(*
SPDX-FileCopyrightText: © 2026 Oleksandr Tiutyk <trofimich@gmail.com>
SPDX-License-Identifier: MIT
License: https://opensource.org/license/mit
*)

(*!
<summary>
Defines a composite activity that waits until the first branch condition becomes TRUE and runs its activity.
</summary>
*)

INTERFACE IWaitAndPickActivity EXTENDS IExclusiveCompositeActivity

(*!
<summary>Appends a condition-activity branch pair and returns its zero-based branch index.</summary>
<description>
Permitted only in PASSIVE_READY. Both condition and activity are required and must not be attached elsewhere.
The standard implementation also rejects duplicate slots, validates fixed workflow association and requires
the parent chain and owning workflow to be PASSIVE_READY before mutation. Child storage remains borrowed.
</description>
<param name="condition">Condition evaluated when polling branches in registration order.</param>
<param name="activity">Activity executed once condition evaluates to TRUE.</param>
*)
METHOD AddBranch : DINT
VAR_INPUT
	condition : ICondition;
	activity : IActivity;
END_VAR
END_METHOD

(*!
<summary>Returns the activity of the currently picked branch, or 0 while waiting or idle.</summary>
*)
{attribute 'monitoring' := 'call'}
PROPERTY CurrentActivity : IActivity
GET
END_GET
END_PROPERTY

(*!
<summary>Returns the zero-based index of the currently picked branch, or -1 while waiting or idle.</summary>
*)
{attribute 'monitoring' := 'call'}
PROPERTY CurrentBranchIndex : DINT
GET
END_GET
END_PROPERTY

END_INTERFACE

(* stored: Version 1.1.0.1
   Itf IWaitAndPickActivity: Id {7c324977-e60a-45fb-9360-b0ea3e5e5a57}
   Method AddBranch: Id {cceb521c-fa78-4662-bb9f-0d9fd6a8e81a}
   Property CurrentActivity: Id {bb402ee2-2866-4ba0-9ad2-a370ad0e4104}
   Get Get: Id {b705ff2e-5341-48ec-ab21-7fbc8de677f7}
   Property CurrentBranchIndex: Id {32f18dd6-a162-4250-9243-ea54bc3d502c}
   Get Get: Id {d27bf5f9-7556-466e-82b0-91ec1d21094c} *)
